// FB_PendantControl with the cover block and the hydraulics block behind it, each in its rig (FB_CoverRig, FB_HydraulicsRig).
// The other blocks the pendant can reference (focus, elevation, azimuth, derotator, telescope) are not connected: the pendant
// must light the error lamp and do nothing for those selections (#16). The test sets the pendant inputs through SetKey(),
// SetSelector(), SetUp() ... and reads the lamps through Lamps() ("x" = lit, order up, down, left, right, error).
// The pendant runs before the blocks in every scan, like in MAIN. StepStart()/nStepScans count the scans from the start of a step.
FUNCTION_BLOCK FB_PendantRig
VAR_INPUT
	stIn		: HalfBROT.ST_PendantIn;
END_VAR
VAR
	fbComm		: FB_NullComm;
	fb			: HalfBROT.FB_PendantControl(comm := fbComm);
	stOut		: HalfBROT.ST_PendantOut;
	cov			: FB_CoverRig;
	hyd			: FB_HydraulicsRig;
	tonStep		: TON;
	nScans		: UDINT;
	nStepScans	: UDINT;
END_VAR

METHOD Scan
nScans := nScans + 1;
nStepScans := nStepScans + 1;
fb(stIn := stIn, fbCovers := cov.fb, fbBrake := hyd.fb, fbHydraulics := hyd.fb, stOut := stOut);
cov.Scan();
hyd.Scan();
tonStep(IN := TRUE, PT := T#1H);
END_METHOD

METHOD SetKey
VAR_INPUT
	bOn	: BOOL;
END_VAR
stIn.bKeySwitch := bOn;
END_METHOD

METHOD SetUp
VAR_INPUT
	bOn	: BOOL;
END_VAR
stIn.bDirectionUp := bOn;
END_METHOD

METHOD SetDown
VAR_INPUT
	bOn	: BOOL;
END_VAR
stIn.bDirectionDown := bOn;
END_METHOD

METHOD SetLeft
VAR_INPUT
	bOn	: BOOL;
END_VAR
stIn.bDirectionLeft := bOn;
END_METHOD

METHOD SetRight
VAR_INPUT
	bOn	: BOOL;
END_VAR
stIn.bDirectionRight := bOn;
END_METHOD

METHOD SetStart
VAR_INPUT
	bOn	: BOOL;
END_VAR
stIn.bStartSwitch := bOn;
END_METHOD

METHOD SetReset
VAR_INPUT
	bOn	: BOOL;
END_VAR
stIn.bResetSwitch := bOn;
END_METHOD

METHOD SetSelector
VAR_INPUT
	nSelector	: INT;
END_VAR
stIn.bBCD0 := (nSelector AND 1) <> 0;
stIn.bBCD2 := (nSelector AND 2) <> 0;
stIn.bBCD4 := (nSelector AND 4) <> 0;
stIn.bBCD8 := (nSelector AND 8) <> 0;
END_METHOD

METHOD SetClearing
VAR_INPUT
	bOn	: BOOL;
END_VAR
hyd.bClearing := bOn;
END_METHOD

METHOD Lamps : STRING(5)
Lamps := '';
IF stOut.bLampUp THEN
	Lamps := CONCAT(Lamps, 'x');
ELSE
	Lamps := CONCAT(Lamps, '-');
END_IF
IF stOut.bLampDown THEN
	Lamps := CONCAT(Lamps, 'x');
ELSE
	Lamps := CONCAT(Lamps, '-');
END_IF
IF stOut.bLampLeft THEN
	Lamps := CONCAT(Lamps, 'x');
ELSE
	Lamps := CONCAT(Lamps, '-');
END_IF
IF stOut.bLampRight THEN
	Lamps := CONCAT(Lamps, 'x');
ELSE
	Lamps := CONCAT(Lamps, '-');
END_IF
IF stOut.bLampError THEN
	Lamps := CONCAT(Lamps, 'x');
ELSE
	Lamps := CONCAT(Lamps, '-');
END_IF
END_METHOD

METHOD State : STRING(100)
State := CONCAT('[sel ', UINT_TO_STRING(fb.Selection));
State := CONCAT(State, CONCAT(' lamps ', Lamps()));
State := CONCAT(State, CONCAT(' open ', cov.OpenOutputs()));
State := CONCAT(State, CONCAT(' close ', cov.CloseOutputs()));
State := CONCAT(State, CONCAT(' pump ', BOOL_TO_STRING(hyd.stOut.bOilPumpEnable)));
State := CONCAT(State, ']');
END_METHOD

METHOD StepStart
tonStep(IN := FALSE, PT := T#1H);
nStepScans := 0;
END_METHOD

METHOD StepTime : BOOL
VAR_INPUT
	tTime	: TIME;
END_VAR
StepTime := tonStep.ET >= tTime;
END_METHOD

END_FUNCTION_BLOCK

(* stored: Version 1.1.0.1, ProductVersion 3.1.4024.15
   POU FB_PendantRig: Id {19e4a2ee-6635-5983-8090-2ff5ba25d08c}, SpecialFunc None
   Method Scan: Id {6e9c1f40-0ef0-559b-8ff1-78659aeeba22}
   Method SetKey: Id {bacc161b-e70c-54fc-9c91-c195e2669dc1}
   Method SetUp: Id {1cf37d19-015c-527d-a70c-c6c1830182e1}
   Method SetDown: Id {559f8eda-7cd6-5ce5-a064-6b29010bc0ca}
   Method SetLeft: Id {db106218-ab9f-5aab-9b03-f800a30a574d}
   Method SetRight: Id {843c2ae9-5ce9-583d-b6f4-3816c74ee7a2}
   Method SetStart: Id {28087647-e35c-5bd7-93b4-f12c3fd6740d}
   Method SetReset: Id {4fb4742d-7569-5d2a-9f60-2d0377a4e72b}
   Method SetSelector: Id {bf6403d8-ee24-529f-8f59-93f59fdaee83}
   Method SetClearing: Id {94eb4b73-5509-5442-894d-135ed913d7c4}
   Method Lamps: Id {8103a3b6-df76-502d-889c-8fa32aba49aa}
   Method State: Id {18dab1ee-83e9-5291-af29-6df26612cc86}
   Method StepStart: Id {5843fba7-9088-53a9-90d6-44acab85be51}
   Method StepTime: Id {6af8c895-718b-574b-9112-e16f110f59e6} *)
